Fanuc KAREL source: KT00746.KL

PROGRAM KT00746
%NOLOCKGROUP
VAR
  ARG: ARRAY[4] OF JOINTPOS
  OUT: BOOLEAN
BEGIN
  OUT = UNINIT(ARG)
END KT00746
